(* PLC project fbd_counter_reset, Anonymous Benchmark Suite 1.0 *)
(* stored: creationDateTime 2026-08-29T00:00:00 *)

PROGRAM drive
  VAR_INPUT
    Reset : BOOL;
    ResetCounterValue : INT;
  END_VAR
  VAR_OUTPUT
    OUT : INT;
  END_VAR
  VAR
    Cnt : INT;
  END_VAR

(* FBD diagram, written out as Structured Text *)
Cnt := SEL(Reset, 1 + Cnt, ResetCounterValue);
OUT := Cnt;
END_PROGRAM

CONFIGURATION Config0
  RESOURCE Res0 ON PLC
    TASK tcyclic(INTERVAL := T#10ms, PRIORITY := 0);
    PROGRAM inst0 WITH tcyclic : drive;
  END_RESOURCE
END_CONFIGURATION
